// TIA Portal V20 export
// export: Created 2026-11-12T11:17:33.8643258Z, ExportSetting WithDefaults, DisplayName Totally Integrated Automation Portal, DisplayVersion V20, DisplayName TIA Portal Openness, DisplayVersion V20, DisplayName TIA Portal Teamcenter Gateway, DisplayVersion V20, DisplayName TIA Portal Version Control Interface, DisplayVersion V20, DisplayName STEP 7 Professional, DisplayVersion V20, DisplayName STEP 7 CFC, DisplayVersion V20, DisplayName STEP 7 Safety, DisplayVersion V20, DisplayName WinCC Basic/Comfort/Advanced, DisplayVersion V20, DisplayName SIMATIC Visualization Architect, DisplayVersion V20, DisplayName WinCC Professional, DisplayVersion V20, DisplayName SIMATIC Visualization Architect, DisplayVersion V20, DisplayName WinCC Unified, DisplayVersion V20, DisplayName SIMATIC Visualization Architect, DisplayVersion V20
VAR_GLOBAL   // PLC tag table "Tabla de variables estándar"
   Entradas_APP AT %I0.0 : "UDT_Entradas_APP";
   Entradas_Basico AT %I1.0 : "UDT_Entradas_Basico";
   Entradas_Stopper AT %I42.0 : "UDT_Entradas_Stopper";
   Salidas_Basico AT %Q1.0 : "UDT_Salidas_Basico";
   Salidas_APP AT %Q0.0 : "UDT_Salidas_APP";
   Entradas_RFID AT %I10.0 : "UDT_Entradas_RFID";
   Salidas_RFID AT %Q10.0 : "UDT_Salidas_RFID";
END_VAR
